(* IEC 61131-3 sources: 2026_Projet_YGO_ExcavatriceDragage/CODE/L_SIMULATION (part 2) *)

(* ---- FB_Sim_WinchElectrical.st ---- *)
(* ═══════════════════════════════════════════════════════════════
   🧪 FB_Sim_WinchElectrical — Composite electrique treuil (charge + couplage)
   ───────────────────────────────────────────────────────────────
   🎯 Role : Calcule le couple resistant reel (charge, benne au sol, couplage
   M1/M2) et pilote FB_Sim_WinchMotor. Transition de charge lissee (evite les
   a-coups de couple/vitesse a la bascule seul<->couple ou charge<->benne au sol).
   📄 Doc metier : DOC/WFLOW/CONTRACTS/PLAN_T317_SIMBENCH_TREUIL_ELECTRIQUE.md
   (registre sequence/interface 2026-09-18 -- pas encore integre a AF_Partie-13)
   🧩 Dependances : FB_Sim_WinchMotor
   ═══════════════════════════════════════════════════════════════ *)
FUNCTION_BLOCK PUBLIC FB_Sim_WinchElectrical
VAR_INPUT
    // === CONTRAT LIGHT ===
    Enable                    : BOOL; // --> [CMD] Autorisation generale FB

    // === COMMANDES ===
    StepCmd                   : INT;  // --> [CMD] Palier resistance rotorique actif (1..5)
    DirectionCmd              : INT := 1; // --> [CMD] Sens (1=Montee, -1=Descente)
    NetworkVoltageAct_V       : REAL := 400.0; // --> [HW] Tension reseau mesuree/simulee

    // === CHARGE ===
    LoadFrac_Ratio            : REAL; // --> [CMD] Taux de charge commande/estime (0..1)
    IsBucketGrounded          : BOOL; // --> [HW] TRUE = benne posee/cable detendu -> charge forcee a 0
        // A cabler sur l'image simulee de M2_TensionedCable_DI (NOT IsBucketGrounded) une fois le
        // stimulus expose en amont (GVL_Simulation) -- interface prete, cablage source en attente.
    LoadTransitionFilter_S    : REAL := 0.5; // --> [CFG] Constante de temps lissage charge (evite a-coup)

    // === COUPLAGE M1/M2 ===
    IsCoupledToPeer           : BOOL; // --> [CMD] TRUE = les deux treuils sont couples (benne commune)
        // A cabler sur l'equivalent simule de CoupledBoth/SyncActive (PRG_04_Treuils_Benne) une fois
        // expose en amont -- interface prete, cablage source en attente (lag 1 cycle accepte).
    PeerTorque_Nm             : REAL; // --> [BUS] Couple moteur de l'autre treuil (cycle precedent)
    PeerSpeed_Rpm             : REAL; // --> [BUS] Vitesse physique de l'autre treuil (cycle precedent)

    // === REGLAGES & CONFIGURATION (relayes a FB_Sim_WinchMotor) ===
    NetworkVoltageNom_V          : REAL := 400.0; // --> [CFG] Tension nominale reseau
    MaxTorque_Nm                 : REAL := 3800.0; // --> [CFG] Cmax decrochage -- SYNTHETIQUE
    SlipAtMaxTorqueBase_Ratio    : REAL := 0.08;   // --> [CFG] gmax palier rotor court-circuite
    RotorResistanceOwn_Ohm       : REAL := 0.08;   // --> [CFG] R2 propre rotor
    Inertia_KgM2                 : REAL := 45.0;   // --> [CFG] Inertie ramenee -- SYNTHETIQUE
    SynchronousSpeed_Rpm         : REAL := 1500.0; // --> [CFG] Vitesse synchronisme
    LoadNominalTorque_Nm         : REAL := 2500.0; // --> [CFG] Couple resistant a pleine charge -- SYNTHETIQUE
    LoadFrictionTorque_Nm        : REAL := 80.0;   // --> [CFG] Frottements residuels a vide -- SYNTHETIQUE
    CoupledPeerGain_Ratio         : REAL := 0.5;   // --> [CFG] Poids de l'effort differentiel du pair en mode couple
    CycleTime_S                  : REAL := 0.01;   // --> [CFG] Pas d'integration
END_VAR
VAR_OUTPUT
    // === CONTRAT LIGHT ===
    Ready                     : BOOL; // <-- [STAT] FB pret

    // === RESULTATS PHYSIQUES (relayes de FB_Sim_WinchMotor) ===
    MotorTorque_Nm            : REAL; // <-- [DIAG] Couple electromagnetique, repere de commande
    ResistiveTorqueAct_Nm     : REAL; // <-- [DIAG] Couple resistant reellement applique (charge+couplage, lisse)
    Slip_Ratio                : REAL; // <-- [DIAG] Glissement, repere de commande
    SpeedAct_Rpm               : REAL; // <-- [DIAG] Vitesse physique reelle signee (+montee/-descente)
    IsStalled                 : BOOL; // <-- [DIAG] Decrochage constate
    IsGeneratorMode            : BOOL; // <-- [DIAG] Mode freinage electrique
END_VAR
VAR
    // === SOUS-INSTANCE FB ===
    Motor                     : FB_Sim_WinchMotor; // * [INST] Couple electromagnetique elementaire

    // === ETAT INTERNE ===
    LoadFracFiltered_Ratio     : REAL; // . [LOC] Taux de charge lisse (PT1)
    LoadFracTarget_Ratio       : REAL; // . [LOC] Cible : 0 si benne au sol, sinon LoadFrac_Ratio
    PeerDifferentialTorque_Nm  : REAL; // . [LOC] Effort differentiel du pair en mode couple
    FilterAlpha_Ratio           : REAL; // . [LOC] Coefficient de lissage du pas courant
END_VAR
VAR CONSTANT
    CST_MinFilterTime_S        : REAL := 0.001;
END_VAR

// === §1 GATE NEUTRALISATION ===
IF NOT Enable THEN
    Ready := FALSE;
    MotorTorque_Nm := 0.0;
    ResistiveTorqueAct_Nm := 0.0;
    Slip_Ratio := 0.0;
    SpeedAct_Rpm := 0.0;
    IsStalled := FALSE;
    IsGeneratorMode := FALSE;
    LoadFracFiltered_Ratio := 0.0;
    RETURN;
END_IF;

// === §2 CHARGE LISSEE (benne au sol force la cible a 0, transition sans a-coup) ===
IF IsBucketGrounded THEN
    LoadFracTarget_Ratio := 0.0;
ELSE
    LoadFracTarget_Ratio := LIMIT(0.0, LoadFrac_Ratio, 1.0);
END_IF;

IF LoadTransitionFilter_S > CST_MinFilterTime_S THEN
    FilterAlpha_Ratio := CycleTime_S / (LoadTransitionFilter_S + CycleTime_S);
ELSE
    FilterAlpha_Ratio := 1.0;
END_IF;
LoadFracFiltered_Ratio := LoadFracFiltered_Ratio
    + FilterAlpha_Ratio * (LoadFracTarget_Ratio - LoadFracFiltered_Ratio);

// === §3 COUPLAGE M1/M2 ===
// En mode couple, la benne lie mecaniquement les deux treuils : un ecart de couple entre pairs
// se traduit en effort differentiel de rattrapage (proportionnel a l'ecart de vitesse), pas en
// deux dynamiques d'inertie totalement independantes qui divergent librement.
IF IsCoupledToPeer THEN
    PeerDifferentialTorque_Nm := CoupledPeerGain_Ratio * (SpeedAct_Rpm - PeerSpeed_Rpm)
        * LoadNominalTorque_Nm / MAX(SynchronousSpeed_Rpm, 1.0);
ELSE
    PeerDifferentialTorque_Nm := 0.0;
END_IF;

// === §4 COUPLE RESISTANT APPLIQUE ===
ResistiveTorqueAct_Nm := LoadFrictionTorque_Nm
    + DirectionCmd * LoadFracFiltered_Ratio * LoadNominalTorque_Nm
    + PeerDifferentialTorque_Nm;

// === §5 MOTEUR ELEMENTAIRE ===
Motor(
    Enable := TRUE,
    StepCmd := StepCmd,
    DirectionCmd := DirectionCmd,
    NetworkVoltageAct_V := NetworkVoltageAct_V,
    ResistiveTorque_Nm := ResistiveTorqueAct_Nm,
    NetworkVoltageNom_V := NetworkVoltageNom_V,
    MaxTorque_Nm := MaxTorque_Nm,
    SlipAtMaxTorqueBase_Ratio := SlipAtMaxTorqueBase_Ratio,
    RotorResistanceOwn_Ohm := RotorResistanceOwn_Ohm,
    Inertia_KgM2 := Inertia_KgM2,
    SynchronousSpeed_Rpm := SynchronousSpeed_Rpm,
    CycleTime_S := CycleTime_S
);

MotorTorque_Nm := Motor.MotorTorque_Nm;
Slip_Ratio := Motor.Slip_Ratio;
SpeedAct_Rpm := Motor.SpeedAct_Rpm;
IsStalled := Motor.IsStalled;
IsGeneratorMode := Motor.IsGeneratorMode;

Ready := TRUE;

(* ---- FB_Sim_WinchMotor.st ---- *)
(* ═══════════════════════════════════════════════════════════════
   🧪 FB_Sim_WinchMotor — Couple electromagnetique moteur treuil (rotor bobine)
   ───────────────────────────────────────────────────────────────
   🎯 Role : Couple (formule de Kloss), glissement bidirectionnel, decrochage
   predictif et mode generatrice pour un treuil M1/M2.
   📄 Doc metier : DOC/WFLOW/CONTRACTS/PLAN_T317_SIMBENCH_TREUIL_ELECTRIQUE.md
   (pas encore integre a AF_Partie-13 -- entree F13.06 a creer lot dedie)
   🧩 Dependances : FB_Sim_KlossTorque
   ═══════════════════════════════════════════════════════════════ *)
FUNCTION_BLOCK PUBLIC FB_Sim_WinchMotor
VAR_INPUT
    // === CONTRAT LIGHT ===
    Enable                    : BOOL; // --> [CMD] Autorisation generale FB (TRUE=Autorise)

    // === COMMANDES ===
    StepCmd                   : INT;  // --> [CMD] Palier resistance rotorique actif (1..5)
    DirectionCmd              : INT := 1; // --> [CMD] Sens (1=Montee, -1=Descente)

    // === MESURES / CHARGE ===
    NetworkVoltageAct_V       : REAL := 400.0; // --> [HW] Tension reseau mesuree/simulee
    ResistiveTorque_Nm        : REAL; // --> [CMD] Couple de charge DEJA projete en repere de
        // commande (N_rel) par l'appelant : positif = s'oppose au mouvement commande, negatif =
        // aide le mouvement (ex. gravite en descente -> peut declencher le mode generatrice).
        // Ce FB ne connait pas le taux de charge/la gravite -- calcul delegue a FB_Sim_WinchElectrical.

    // === REGLAGES & CONFIGURATION ===
    NetworkVoltageNom_V          : REAL := 400.0; // --> [CFG] Tension nominale reseau
    MaxTorque_Nm                 : REAL := 3800.0; // --> [CFG] Cmax decrochage -- SYNTHETIQUE
    SlipAtMaxTorqueBase_Ratio    : REAL := 0.08;   // --> [CFG] gmax au palier rotor court-circuite
        // (resistance externe nulle) -- SYNTHETIQUE. Sert de base a la mise a l'echelle par palier.
    RotorResistanceOwn_Ohm       : REAL := 0.08;   // --> [CFG] R2 propre rotor (palier court-circuite)
    Inertia_KgM2                 : REAL := 45.0;   // --> [CFG] Inertie ramenee -- SYNTHETIQUE
    SynchronousSpeed_Rpm         : REAL := 1500.0; // --> [CFG] Vitesse synchronisme
    CycleTime_S                  : REAL := 0.01;   // --> [CFG] Pas d'integration
END_VAR
VAR_OUTPUT
    // === CONTRAT LIGHT ===
    Ready                     : BOOL; // <-- [STAT] FB pret

    // === RESULTATS PHYSIQUES ===
    MotorTorque_Nm            : REAL; // <-- [DIAG] Couple electromagnetique, repere de commande
    Slip_Ratio                : REAL; // <-- [DIAG] Glissement, repere de commande
    SpeedAct_Rpm               : REAL; // <-- [DIAG] Vitesse physique reelle signee (+montee/-descente)
    IsStalled                 : BOOL; // <-- [DIAG] Decrochage constate (jamais reinitialise)
    IsGeneratorMode            : BOOL; // <-- [DIAG] Couple oppose au sens de commande (freinage)
END_VAR
VAR
    // === SOUS-INSTANCES FB ===
    KlossRunning               : FB_Sim_KlossTorque; // * [INST] Couple regime etabli
    KlossLockedRotor           : FB_Sim_KlossTorque; // * [INST] Couple test decrochage (g=1)

    // === ETAT INTERNE ===
    SpeedRel_RadPerS           : REAL; // . [LOC] Vitesse en repere de commande (N_rel)
    SynchronousSpeed_RadPerS   : REAL; // . [LOC] Vitesse synchronisme, rad/s
    SlipAtMaxTorqueStep_Ratio  : REAL; // . [LOC] gmax au palier courant
    SlipEff_Ratio               : REAL; // . [LOC] Glissement protege division par zero
    VoltageRatio2               : REAL; // . [LOC] (U_act/U_nom)^2
    Stalled                    : BOOL; // . [LOC] Etat instantane, peut se relever

    // === ENTREES BORNEES (SECURISE DIVISIONS) ===
    InertiaSafe_KgM2            : REAL; // . [LOC] Inertia_KgM2 bornee > 0
    RotorResistanceOwnSafe_Ohm  : REAL; // . [LOC] RotorResistanceOwn_Ohm bornee > 0
    SlipAtMaxTorqueBaseSafe_Ratio : REAL; // . [LOC] SlipAtMaxTorqueBase_Ratio bornee > 0
    NetworkVoltageNomSafe_V     : REAL; // . [LOC] NetworkVoltageNom_V bornee > 0
    StepCmdSafe                : INT;  // . [LOC] StepCmd borne [1..5]
END_VAR
VAR CONSTANT
    CST_StepCount              : INT := 5;
    CST_RotorExtResistanceStep_Ohm : ARRAY[1..5] OF REAL := [3.6, 1.9, 0.9, 0.35, 0.0];
        // palier 1 = resistance max (demarrage), palier 5 = rotor court-circuite -- SYNTHETIQUE
        // (indexation/valeurs propres au ST, pas un portage 1:1 du prototype Python 4 gradins)
    CST_MinSlip_Ratio          : REAL := 0.0001;
    CST_MinDenominator         : REAL := 0.001; // plancher generique config sensible (division)
    CST_StallSpeedThreshold_Rpm : REAL := 28.0; // ~3 rad/s, "quasi arrete"
END_VAR

// === §1 GATE NEUTRALISATION ===
IF NOT Enable THEN
    Ready := FALSE;
    MotorTorque_Nm := 0.0;
    Slip_Ratio := 0.0;
    SpeedAct_Rpm := 0.0;
    IsStalled := FALSE;
    IsGeneratorMode := FALSE;
    SpeedRel_RadPerS := 0.0;
    RETURN;
END_IF;

StepCmdSafe := LIMIT(1, StepCmd, CST_StepCount);
IF StepCmdSafe <> StepCmd THEN
    Ready := FALSE;
    RETURN;
END_IF;
IF (DirectionCmd <> 1) AND (DirectionCmd <> -1) THEN
    Ready := FALSE;
    RETURN;
END_IF;

// Bornage systematique des entrees de config sensibles (denominateurs) -- CODE_QUALITY_STANDARDS §6
InertiaSafe_KgM2 := MAX(CST_MinDenominator, Inertia_KgM2);
RotorResistanceOwnSafe_Ohm := MAX(CST_MinDenominator, RotorResistanceOwn_Ohm);
SlipAtMaxTorqueBaseSafe_Ratio := MAX(CST_MinDenominator, SlipAtMaxTorqueBase_Ratio);
NetworkVoltageNomSafe_V := MAX(1.0, NetworkVoltageNom_V);

// === §2 GLISSEMENT ET COUPLE (FORMULE DE KLOSS) ===
SynchronousSpeed_RadPerS := SynchronousSpeed_Rpm * 2.0 * 3.14159265 / 60.0;

// gmax(palier) = gmax_base * R2_total(palier) / R2_rotor_propre -- ajouter de la resistance
// externe deplace le glissement au couple max vers 1 (couple demarrage), sans changer Cmax.
// gmax_base = gmax au palier rotor court-circuite (resistance externe nulle).
SlipAtMaxTorqueStep_Ratio := SlipAtMaxTorqueBaseSafe_Ratio
    * (RotorResistanceOwnSafe_Ohm + CST_RotorExtResistanceStep_Ohm[StepCmdSafe])
    / RotorResistanceOwnSafe_Ohm;

// Glissement en repere de commande (N_rel) : peut etre negatif (survitesse -> freinage
// generateur). SpeedRel_RadPerS reste dans ce repere ; SpeedAct_Rpm restitue le signe physique.
Slip_Ratio := 1.0 - SpeedRel_RadPerS / SynchronousSpeed_RadPerS;

IF ABS(Slip_Ratio) < CST_MinSlip_Ratio THEN
    IF Slip_Ratio >= 0.0 THEN
        SlipEff_Ratio := CST_MinSlip_Ratio;
    ELSE
        SlipEff_Ratio := -CST_MinSlip_Ratio;
    END_IF;
ELSE
    SlipEff_Ratio := Slip_Ratio;
END_IF;

VoltageRatio2 := (NetworkVoltageAct_V / NetworkVoltageNomSafe_V) * (NetworkVoltageAct_V / NetworkVoltageNomSafe_V);

KlossRunning(
    Enable := TRUE,
    MaxTorque_Nm := MaxTorque_Nm,
    Slip_Ratio := SlipEff_Ratio,
    SlipAtMaxTorque_Ratio := SlipAtMaxTorqueStep_Ratio,
    VoltageRatio2 := VoltageRatio2);
MotorTorque_Nm := KlossRunning.Torque_Nm;

// === §3 DYNAMIQUE MECANIQUE ===
// Pas de saturation basse : SpeedRel_RadPerS peut devenir negatif (glissement arriere sous
// surcharge) ou depasser le synchronisme (regime generateur).
SpeedRel_RadPerS := SpeedRel_RadPerS
    + (MotorTorque_Nm - ResistiveTorque_Nm) / InertiaSafe_KgM2 * CycleTime_S;

SpeedAct_Rpm := SpeedRel_RadPerS * DirectionCmd * 60.0 / (2.0 * 3.14159265);

// === §4 DECROCHAGE PREDICTIF ===
// Au palier courant, couple disponible a glissement bloque (g=1) < couple resistant, ET
// vitesse quasi nulle -- prediction "ce palier peut-il tenir la charge depuis l'arret ?",
// pas une mesure d'arret reel.
IF ABS(SpeedAct_Rpm) < CST_StallSpeedThreshold_Rpm THEN
    KlossLockedRotor(
        Enable := TRUE,
        MaxTorque_Nm := MaxTorque_Nm,
        Slip_Ratio := 1.0,
        SlipAtMaxTorque_Ratio := SlipAtMaxTorqueStep_Ratio,
        VoltageRatio2 := VoltageRatio2);
    Stalled := KlossLockedRotor.Torque_Nm < ResistiveTorque_Nm;
    IF Stalled THEN
        IsStalled := TRUE;
    END_IF;
ELSE
    Stalled := FALSE;
END_IF;

IsGeneratorMode := MotorTorque_Nm < 0.0;

Ready := TRUE;

(* ---- FB_SimBench.st ---- *)
(* ═══════════════════════════════════════════════════════════════
   🧪 FB_SimBench — Enveloppe unique de simulation pour banc d'essai
   ───────────────────────────────────────────────────────────────
   📄 Doc métier : DOC/AF/AF_Partie-13_Fonction_Simulation_v2.5.md

   🎯 Rôle : Compose les blocs de modèle de simulation :
      - FB_Sim_Encoder (instM1, instM2)
      - FB_Sim_Translation (instTranslation)
      - FB_Sim_Joystick (instJoystick)
      - FB_Sim_Safety (instSafety)

   🔒 Brique réduite : 0 lecture de variable globale en interne.
      Toutes les entrées (commandes, stimuli, HwReal) sont passées en paramètres.

   🔴 RÈGLES SÉCURITÉ ET POLARITÉ :
      - Modèle frein M1/M2/M3 : M1_BrakeIsOpen_DI := M1_BrakeCmd (1 = OUVERT).
        Ne JAMAIS faire NOT BrakeCmd !
      - Retours contacteurs M1/M2 : 1 = tous retombés (TRUE quand RelayFwd=0 et RelayRev=0).
   ═══════════════════════════════════════════════════════════════ *)

FUNCTION_BLOCK PUBLIC FB_SimBench
VAR_INPUT
    Enable                     : BOOL;             (* --> [CMD] Activation globale (GVL_Simulation.SimulationModeActive) *)
    OperatorSourceActive       : BOOL := TRUE;      (* --> [CMD] Source operateur simulee effectivement selectionnee *)

    // ── Commandes issues de l'automate (Scan N-1 / PRG_07 / PRG_10) ──────────
    M1_RelayFwd                : BOOL;   (* --> [CMD] Sens avant M1 *)
    M1_RelayRev                : BOOL;   (* --> [CMD] Sens arrière M1 *)
    // Les 4 contacteurs de palier participent au retour unique
    // « tous contacteurs retombés » — sans eux, le modèle annonce l'arrêt alors qu'un
    // palier est encore engagé (fausse condition d'armement Méca A).
    M1_SpeedContactor_1        : BOOL;   (* --> [HW] Contacteur palier 1 M1 *)
    M1_SpeedContactor_2        : BOOL;   (* --> [HW] Contacteur palier 2 M1 *)
    M1_SpeedContactor_3        : BOOL;   (* --> [HW] Contacteur palier 3 M1 *)
    M1_SpeedContactor_4        : BOOL;   (* --> [HW] Contacteur palier 4 M1 *)
    M1_SpeedCmd_Pct            : REAL;   (* --> [CMD] Consigne vitesse M1 *)
    M1_StepNumber              : INT;    (* --> [CMD] Palier vitesse courant M1 (1..5) *)
    M1_PresetTriggerCmd        : WORD;   (* --> [CMD] Trigger preset M1 *)
    M1_PresetValueOut          : UDINT;   (* --> [CFG] Valeur preset M1 *)
    M1_BrakeCmd                : BOOL;             (* --> [CMD] TRUE = commande desserrage frein M1 *)

    M2_RelayFwd                : BOOL;   (* --> [CMD] Sens avant M2 *)
    M2_RelayRev                : BOOL;   (* --> [CMD] Sens arrière M2 *)
    M2_SpeedContactor_1        : BOOL;   (* --> [HW] Idem M1, voir ci-dessus *)
    M2_SpeedContactor_2        : BOOL;   (* --> [HW] Contacteur palier 2 M2 *)
    M2_SpeedContactor_3        : BOOL;   (* --> [HW] Contacteur palier 3 M2 *)
    M2_SpeedContactor_4        : BOOL;   (* --> [HW] Contacteur palier 4 M2 *)
    M2_SpeedCmd_Pct            : REAL;   (* --> [CMD] Consigne vitesse M2 *)
    M2_StepNumber              : INT;    (* --> [CMD] Palier vitesse courant M2 (1..5) *)
    M2_PresetTriggerCmd        : WORD;   (* --> [CMD] Trigger preset M2 *)
    M2_PresetValueOut          : UDINT;   (* --> [CFG] Valeur preset M2 *)
    M2_BrakeCmd                : BOOL;             (* --> [CMD] TRUE = commande desserrage frein M2 *)

    M3_ReqTremie               : BOOL;             (* --> [CMD] Demande explicite vers Trémie *)
    M3_ReqMaintenance          : BOOL;             (* --> [CMD] Demande explicite vers Maintenance *)
    M3_SpeedCmd_Pct            : REAL;   (* --> [CMD] Consigne vitesse M3 *)
    (* T301/L1 — SOURCE UNIQUE : reglages machine M3 lus par PRG_02 (le banc n'a plus de positions en dur) *)
    M3_PosTremie_M             : REAL := 0.0;   (* --> [CFG] Position capteur Tremie (GVL_PERSISTENT) *)
    M3_PosPV_M                 : REAL := 1.5;   (* --> [CFG] Position capteur PV (GVL_PERSISTENT) *)
    M3_PosP2_M                 : REAL := 3.5;   (* --> [CFG] Position capteur P2 (GVL_PERSISTENT) *)
    M3_PosP1_M                 : REAL := 5.0;   (* --> [CFG] Position capteur P1 (GVL_PERSISTENT) *)
    M3_PosMaintenance_M        : REAL := 10.0;  (* --> [CFG] Position capteur Maintenance (GVL_PERSISTENT) *)
    M3_OdometryGain            : REAL := 0.02;  (* --> [CFG] Gain effectif de l'estimateur machine, m/(Hz.s) (PRG_05) *)
    M3_EstimatedPos_M          : REAL;          (* --> [DIAG] Position calculee par le programme (PRG_05), pour l'ecart observe *)
    M3_BrakeCmd                : BOOL;             (* --> [CMD] TRUE = commande desserrage frein M3 *)

    PowerKeepAlive_A           : BOOL;             (* --> [SAFE] TRUE = relais A maintenu sagement par le PLC *)
    PowerKeepAlive_B           : BOOL;             (* --> [SAFE] TRUE = relais B maintenu sagement par le PLC *)
    EmergencyArming_RQ         : BOOL;             (* --> [CMD] Impulsion de réarmement puissance *)
    TestCutActive              : BOOL;             (* --> [SAFE] Test de redondance AU en cours (canal A ou B coupé) *)
    PowerCutOffRequest         : BOOL;             (* --> [SAFE] Requête coupure métier (TRUE = arrêt d'urgence) *)
    SimChainOkBit              : BOOL;             (* --> [TST] Bit opérateur : TRUE = simuler chaîne AU fermée *)
    SimPhaseRotationOkBit      : BOOL;             (* --> [TST] Bit opérateur : TRUE = phases réseau OK ; FALSE = défaut rotation de phases *)

    // ── Stimuli & Paramètres de banc ─────────────────────────────────────────
    SimEncoderSpeedFactor      : REAL := 1.0;   (* --> [CFG] Facteur vitesse codeur *)
    SimBucketSpeedFactor       : REAL := 1.0;   (* --> [CFG] Facteur vitesse manoeuvre benne seule (non persistant) *)
    SimTopPositionActive       : BOOL := FALSE; (* --> [TST] Injection manuelle capteur haut actif (essai ciblé) *)
    SimSyncDeviationInjectM1   : BOOL := FALSE;   (* --> [TST] Injection écart synchro M1 *)
    SimSyncDeviationInjectM2   : BOOL := FALSE;   (* --> [TST] Injection écart synchro M2 *)
    SimSyncDeviationOffset_M   : REAL := 0.5;   (* --> [TST] Offset écart synchro *)
    SimM2CoupledDescentModelActive : BOOL := TRUE; (* --> [CFG] M2 calculé depuis M1 en descente BOTH *)
    SimM2CoupledDescentFactor  : REAL := 0.9333; (* --> [CFG] Ratio déplacement M2/M1 mesuré: 0,6m d'écart sur 9m *)
    SimWinchSpeedReportTauS    : REAL := 0.0;    (* --> [CFG][SYNTHETIQUE] Tau 1er ordre retour vitesse rapportee M1/M2, s. 0.0 = saut instantane (comportement historique). *)
    SimWinchBrakeOpenDelayS    : REAL := 0.0;    (* --> [CFG][SYNTHETIQUE] Delai electrique/meca ouverture frein M1/M2 apres BrakeCmd=TRUE, s. 0.0 = instantane (comportement historique). *)
    SimWinchBrakeCloseDelayS   : REAL := 0.0;    (* --> [CFG][SYNTHETIQUE] Delai electrique/meca fermeture frein M1/M2 apres BrakeCmd=FALSE, s. 0.0 = instantane (comportement historique). *)
    SimWinchDynamicsActive     : BOOL := FALSE;  (* --> [CFG] TRUE = applique tau et delais treuils ; FALSE = profil simple historique *)

    // T317 exploratoire -- charge/couplage electrique treuil (interface prete, defaut = comportement
    // historique inchange tant que non cablee sur un vrai signal amont, cf. registre PLAN_T317).
    SimWinchLoadFrac_Ratio     : REAL := 0.0;    (* --> [CFG][SYNTHETIQUE] Taux de charge M1/M2, 0=a vide *)
    SimWinchCoupledActive      : BOOL := FALSE;  (* --> [TST] M1/M2 couples -- en attente cablage CoupledBoth reel *)
    SimWinchElectricalDiagnosticsActive : BOOL := FALSE; (* --> [CFG] TRUE = publie diagnostic electrique treuils, sans action safety *)
    SimM2TensionedCableFaultInject : BOOL := FALSE; (* --> [TST] TRUE = injecte capteur cable non tendu M2 *)

    SimM3SensorsWordOverrideActive : BOOL := FALSE;   (* --> [TST] Override mot capteurs M3 *)
    SimM3SensorsWord               : BYTE := 16#07;   (* --> [TST] Mot capteurs M3 forcé *)
    SimM3SensorIntermittenceActive  : BOOL := FALSE;   (* --> [TST] Episode perte/reprise DI M3 *)
    SimM3SensorStabilizationS       : REAL := 1.0;     (* --> [CFG] Duree episode capteur M3, s *)
    SimM3SensorElectricalDelayS     : REAL := 0.01;    (* --> [CFG] Delai electrique capteur M3, s *)
    SimM3SensorIntermittencePeriodS : REAL := 0.12;    (* --> [CFG] Periode des bascules episode, s *)
    SimM3SensorHysteresis_M         : REAL := 0.02;    (* --> [CFG] Hysteresis seuils capteurs M3, m *)
    SimM3SensorLoadAngleTriggerRad  : REAL := 0.01;    (* --> [CFG] Angle charge minimal episode, rad *)
    SimM3SensorScenarioSeed         : UDINT := 3001;   (* --> [CFG] Graine episode capteurs M3 *)
    SimM3SensorBlipTransitions      : UDINT := 0;      (* --> [TST] Excursions electriques courtes par front (0 = profil ~1 s historique seul) *)
    SimM3SensorBlipDurationS        : REAL := 0.2;     (* --> [CFG] Largeur d'une excursion du blip court, s *)
    // FAUTE explicite frein M3 — defaut FALSE : reproduit le defaut terrain « frein ferme
    // alors que le variateur retourne encore 10,00 Hz » (trace 2026-09-04, 26,437 s, ErrorId=64).
    SimM3BrakeFaultCloseWhileRunning : BOOL := FALSE;  (* --> [TST] TRUE = force la fermeture frein M3 hors vitesse nulle *)
    SimM3BrakeFaultCloseDelayS       : REAL := 0.0;    (* --> [CFG] Delai avant application de la faute frein M3, s *)
    SimM3BrakePhysicalActive         : BOOL := TRUE;   (* --> [CFG] L3 : frein M3 a manque de courant reel (FALSE = historique) *)
    SimM3BrakeDecel_Mps2             : REAL := 2.0;    (* --> [CFG][HYPOTHESE] Deceleration chariot frein serre, m/s2 *)
    SimM3CartFreeActive              : BOOL := TRUE;   (* --> [CFG] L4 : chariot libre frein ouvert + variateur sans couple *)
    SimM3LoadMassRatio               : REAL := 0.5;    (* --> [CFG][HYPOTHESE] Masse benne / masse totale *)
    SimM3RollingFriction_Mps2        : REAL := 0.1;    (* --> [CFG][HYPOTHESE] Frottement de roulement, m/s2 *)
    SimM3Slope_Mps2                  : REAL := 0.0;    (* --> [CFG][HYPOTHESE] Pente, m/s2 (+ vers Maintenance) *)
    SimM3SensorCamDropoutActive      : BOOL := TRUE;   (* --> [CFG] L5 : came capteurs vu -> perdu -> retrouve -> fixe *)
    SimM3SensorCamDropoutStart_M     : REAL := 0.02;   (* --> [CFG][HYPOTHESE] Debut de la zone perdue apres la cote, m *)
    SimM3SensorCamDropoutWidth_M     : REAL := 0.04;   (* --> [CFG][HYPOTHESE] Largeur de la zone perdue, m *)
    // BUTEE MECANIQUE M3 — recul borne apres arret serre (C5). 0.0 = comportement historique
    // (position ET vitesse figees a la butee, decision de review tracee). > 0 autorise la
    // reaction de charge a ressortir le chariot de la zone capteur. SYNTHETIQUE, non calibre.
    SimM3EndStopRecoilMax_M          : REAL := 0.0;    (* --> [CFG][SYNTHETIQUE] Recul borne a la butee M3, m *)
    SimM3EndStopMargin_M             : REAL := 0.5;    (* --> [CFG] Distance capteur extreme -> butee mecanique M3, m *)
    SimM3LoadReactionGain_Mps2       : REAL := 0.20;   (* --> [CFG][SYNTHETIQUE] Gain de reaction de charge M3, m/s2 *)
    // ACCELERATION DU BANC M3 : chariot ET frequence retournee x facteur (1..5), estimation coherente.
    // Volontairement NON cable par PRG_02 : se regle en ligne sur l'instance (instSimBench.SimM3SpeedFactor).
    SimM3SpeedFactor                 : REAL := 1.0;    (* --> [TST] Facteur de vitesse du banc M3, 1,0 = dynamique reelle *)

    SimJoystickLeft_Rev_TREMIE_Active  : BOOL := FALSE;   (* --> [TST] Bouton joystick gauche *)
    SimJoystickRight_Fwd_MAINT_Active  : BOOL := FALSE;   (* --> [TST] Bouton joystick droite *)
    SimJoystickFwd_Up_Close_Active     : BOOL := FALSE;   (* --> [TST] Bouton joystick avant *)
    SimJoystickRev_Down_Open_Active    : BOOL := FALSE;   (* --> [TST] Bouton joystick arrière *)
    SimJoystickRawX                    : INT := 5000;   (* --> [TST] Valeur brute X *)
    SimJoystickRawY                    : INT := 5000;   (* --> [TST] Valeur brute Y *)
    SimJoystickRawButton               : BOOL := FALSE;   (* --> [TST] Bouton homme-mort *)
    SimJoystickOvershoot_Active        : BOOL := FALSE;   (* --> [TST] Dépassement de montée au-delà de 100% (défaut capteur hors plage) *)
    SimJoystickBagotement_Active       : BOOL := FALSE;   (* --> [TST] Bagotement au relâchement (petit balancement autour du neutre) *)

    SimKoboldContactValue      : BOOL := FALSE;   (* --> [TST] Contact fond Kobold *)
    SimKoboldAutoModeActive    : BOOL := FALSE;   (* --> [CFG] Kobold positionnel automatique armé *)
    SimKoboldAutoDepth_M       : REAL := -15.0;   (* --> [CFG] Fond Kobold signé *)
    SimKoboldPowerUpTime       : TIME := T#50ms;  (* --> [CFG] Temps de réponse sonde *)
    SimKoboldCoast_M           : REAL := 1.0;     (* --> [CFG] Compatibilité interface ; dynamique historique utilisée *)
    KoboldMeasureEnable        : BOOL := FALSE;   (* --> [CMD] Alimentation Kobold effectivement arbitrée *)
    M1_CablePos_M              : REAL := 0.0;     (* --> [HW] Position M1 signée, référence homing effective *)
    BtnEmergencyStop           : BOOL := FALSE;    (* --> [TST] Simulation appui coup-de-poing AU *)

    // ── Rattrapage mécanique M1/M2 (reprise de jeu en mouvement couplé) ──
    SimWinchCouplingModelActive : BOOL := TRUE;    (* --> [CFG] TRUE = rattrapage mécanique modélisé au banc *)
    SimBucketJamActive          : BOOL := FALSE;   (* --> [TST] TRUE = mâchoires bloquées (objet coincé) *)
    WinchesHomed                : BOOL := TRUE;    (* --> [HW] TRUE = M1 et M2 references (butee meca benne inactive avant homing) *)
    M2_CablePos_M               : REAL := 0.0;     (* --> [HW] Position M2 recalée (m), issue de la même chaîne que le métier *)
    BucketOffsetCloseM          : REAL := 15.0;    (* --> [CFG] Butée mécanique benne FERMÉE (m, écart M2-M1) *)
    BucketCoherenceLimitM       : REAL := 1.0;     (* --> [CFG] Demi-largeur de la bande franc ouvert/fermé (m) *)
    BucketOffsetOpen_M          : REAL := 0.0;     (* --> [CFG] Butée mécanique benne OUVERTE (m, écart M2-M1) *)
    BucketOpenAnticipation_M    : REAL := 1.3;     (* --> [CFG] Anticipation arrêt ouverture benne (m) *)
    BucketAx15bOpenActive       : BOOL := FALSE;   (* --> [CMD] Étape AX15B active *)

    // ── Image réelle fallback ────────────────────────────────────────────────
    HwReal                     : ST_HardwareImage;   (* --> [HW] Image réelle fallback *)
END_VAR

VAR_OUTPUT
    (* Sorties d'état du profil AF_Partie-03 §2.
       En LD, CODESYS réserve la PREMIÈRE broche de sortie au flux du rung :
       `Ready` n'y porte jamais d'expression, les broches suivantes oui. *)
    Ready                      : BOOL;             (* <-- [STAT] TRUE = banc prêt (Enable actif, modèles à jour) *)
    Busy                       : BOOL;             (* <-- [STAT] TRUE = cycle de simulation en cours *)
    Done                       : BOOL;             (* <-- [STAT] TRUE = images de simulation publiées ce scan *)

    Winch                      : ST_HwWinch;   (* <-- [DIAG] Image treuils simulée *)
    Translation                : ST_HwTranslation;   (* <-- [DIAG] Image translation simulée *)
    Operator                   : ST_HwOperator;   (* <-- [DIAG] Image opérateur simulée *)
    Machine                    : ST_HwMachine;   (* <-- [DIAG] Image machine simulée *)

    // T317 exploratoire -- modele electrique treuil, diagnostic seul, non consomme par le metier.
    // Charge appliquee = LoadFrictionTorque_Nm + taux x LoadNominalTorque_Nm (FB_Sim_WinchElectrical) ;
    // le taux de charge n'est pas encore cable sur un signal amont (registre PLAN_T317).
    MotorTorqueM1_Nm           : REAL;   (* <-- [DIAG] T317 -- Couple electromagnetique simule M1 *)
    MotorTorqueM2_Nm           : REAL;   (* <-- [DIAG] T317 -- Couple electromagnetique simule M2 *)
    MotorIsStalledM1           : BOOL;   (* <-- [DIAG] T317 -- Decrochage predictif simule M1 *)
    MotorIsStalledM2           : BOOL;   (* <-- [DIAG] T317 -- Decrochage predictif simule M2 *)

    // Rattrapage mecanique M1/M2 -- diagnostic seul (aucun consommateur metier).
    WinchCouplingActive        : BOOL;   (* <-- [DIAG] Rattrapage applique ce scan *)
    WinchCouplingCorrectionPts : DINT;   (* <-- [DIAG] Correction appliquee a l'image M2 (points codeur) *)

    // Faute frein M3 -- diagnostic seul : confirme que la branche de faute est bien appliquee.
    M3BrakeFaultCloseActive    : BOOL;   (* <-- [DIAG] Faute frein M3 effectivement appliquee ce scan *)
    // Blip court capteurs M3 -- diagnostic seul : observable sur trace pendant un episode court.
    M3SensorBlipActive         : BOOL;   (* <-- [DIAG] Un capteur M3 publie une excursion courte *)
    (* L2 — observation M3 (lecture seule, aucun effet sur le pilotage) *)
    M3ObsPositionTrue_M        : REAL;   (* <-- [DIAG] Position vraie du chariot simule (m) *)
    M3ObsPositionError_M       : REAL;   (* <-- [DIAG] Position vraie - position calculee par le programme (m) *)
    M3ObsOvershootLast_M       : REAL;   (* <-- [DIAG] Distance roulee apres le 1er front du dernier capteur d'arret (m) *)
    M3ObsOvershootSensorId     : INT;    (* <-- [DIAG] 1 = Tremie, 3 = P1, 5 = Maintenance *)
    M3ObsEndStopHitCount       : UDINT;  (* <-- [DIAG] Chocs en butee mecanique *)
    M3ObsEndStopImpactSpeed_Mps : REAL;  (* <-- [DIAG] Vitesse au dernier choc en butee (m/s) *)
    M3ObsBrakeClosedMovingCount : UDINT; (* <-- [DIAG] Fermetures du frein chariot en mouvement *)
    M3ObsCartFree              : BOOL;   (* <-- [DIAG] L4 : chariot libre (frein ouvert, variateur sans couple) *)
    M3ObsFreeRollLast_M        : REAL;   (* <-- [DIAG] L4 : distance du dernier episode libre (m) *)
END_VAR

VAR_IN_OUT
    // 🔒 LECTURE SEULE pour le banc : ces mémoires appartiennent au modèle codeur. Le banc les lit
    //    pour piloter ses modèles et ne les écrit JAMAIS — pas même pour « initialiser » une mémoire
    //    lue à 0 (un 0 est un point de passage légitime du comptage signé, jamais une mémoire vierge).
    RawPosM1                   : UDINT;            (* <-> [BUS] Mémoire _SimEncoderRawPosM1 dans GVL_PERSISTENT *)
    RawPosM2                   : UDINT;            (* <-> [BUS] Mémoire _SimEncoderRawPosM2 dans GVL_PERSISTENT *)
END_VAR

VAR CONSTANT
    // T301/L1 : l'ancienne echelle en dur CST_M3FullTravelTimeS (37,5 s) est SUPPRIMEE — le banc
    // recoit positions + gain effectif de la machine (M3_Pos*_M, M3_OdometryGain). Gate G518.
    // Maximum variateur M3 : DOIT egaler GVL_PERSISTENT._TranslationMaxFreq_Hz (PRG_02 envoie f/50 x 100).
    // Constante locale (L_SIMULATION ne lit pas GVL_PERSISTENT) ; egalite verifiee par G518.
    CST_M3MaxFreq_Hz            : REAL := 50.0;
    CST_SimBenchCycleTimeS      : REAL := 0.010; // Période tâche PLC (s) — MainTask 10 ms
    // Rattrapage mécanique M1/M2 — valeurs ESTIMÉES (voir REGISTRE_VALEURS_TREUIL_STATUTS_v1.0.md)
    CST_SimWinchCouplingTauS    : REAL := 1.0;   // [HYPOTHESE] Constante de temps du rattrapage (s)
    CST_SimWinchCouplingStepMax_M : REAL := 0.02; // [HYPOTHESE] Borne de pente par scan (= 2,0 m/s x 0,010 s)
    CST_SimWinchCouplingPtsPerM : REAL := 4096.0; // Points codeur par mètre (8192 pts/tour / 2,0 m/tour)
    CST_SimBucketJamLoadFrac_Ratio : REAL := 1.0; // [HYPOTHESE] Charge forcée quand les mâchoires sont bloquées
END_VAR

VAR
    // Modèles sous-jacents
    instSimEncoderM1           : FB_Sim_Encoder;   (* * [INST] Modèle codeur M1 *)
    instSimEncoderM2           : FB_Sim_Encoder;   (* * [INST] Modèle codeur M2 *)
    instSimTranslation         : FB_Sim_Translation;   (* * [INST] Modèle translation M3 *)
    instSimJoystick            : FB_Sim_Joystick;   (* * [INST] Modèle joystick *)
    instSimSafety              : FB_Sim_Safety;   (* * [INST] Modèle sécurité *)
    instWinchElectricalM1      : FB_Sim_WinchElectrical;   (* * [INST] T317 exploratoire -- electrique+charge M1 *)
    instWinchElectricalM2      : FB_Sim_WinchElectrical;   (* * [INST] T317 exploratoire -- electrique+charge M2 *)
    PeerTorqueM1Prev_Nm        : REAL;   (* . [LOC] T317 -- couple M1 cycle precedent, pour M2 couple *)
    PeerTorqueM2Prev_Nm        : REAL;   (* . [LOC] T317 -- couple M2 cycle precedent, pour M1 couple *)
    PeerSpeedM1Prev_Rpm        : REAL;   (* . [LOC] T317 -- vitesse M1 cycle precedent, pour M2 couple *)
    PeerSpeedM2Prev_Rpm        : REAL;   (* . [LOC] T317 -- vitesse M2 cycle precedent, pour M1 couple *)
    KoboldBottomTouchPrev_DI   : BOOL;   (* . [LOC] T317 -- Machine.M1_M2_KoboldBottomTouch_DI cycle precedent (benne au sol) *)

    // Calculs internes
    M1_PresetCmd               : BOOL;   (* . [LOC] Trigger preset M1 *)
    M2_PresetCmd               : BOOL;   (* . [LOC] Trigger preset M2 *)
    M1_OffsetPts               : DINT;   (* . [LOC] Offset synchro M1 *)
    M2_OffsetPts               : DINT;   (* . [LOC] Offset synchro M2 *)

    M3_RelayFwd                : BOOL;   (* . [LOC] Sens avant M3 *)
    M3_RelayRev                : BOOL;   (* . [LOC] Sens arrière M3 *)

    SimJoystickManualNeutral : BOOL; (* . [LOC] Axes manuels au neutre nominal *)
    SimJoystickGesturePermit : BOOL; (* . [LOC] Aucune injection manuelle concurrente au geste *)

    M3_ActualFreqHz            : UINT;   (* . [LOC] Fréquence simulée M3 *)
    M3_StatusWordSim           : WORD;   (* . [LOC] StatusWord simulé M3 *)

    // Roulis dynamique avec dispersion pseudo-aléatoire (±0.1m autour de l'anticipation)
    M2_RelayFwdPrev            : BOOL;   (* . [LOC] Mémoire relais Fwd N-1 *)
    M2_RelayRevPrev            : BOOL;   (* . [LOC] Mémoire relais Rev N-1 *)
    RandomSeed                 : UDINT := 123456789; (* . [LOC] Générateur LCG pseudo-aléatoire *)
    M2_EffectiveCoastM         : REAL := 1.30;       (* . [LOC] Distance de roulis M2 courante *)
    M2EffectiveCoastDistance_M : REAL;               (* . [LOC] Distance appliquée au codeur M2 *)
    M2AutoOpenCoastArmed       : BOOL;               (* . [LOC] Fin d'ouverture automatique à simuler *)
    M2OpenDistanceRemaining_M  : REAL;               (* . [LOC] Distance restante à la butée ouverte *)
    M2OpenStopThreshold_M     : REAL;               (* . [LOC] Seuil avec avance d'un scan d'acquisition *)
    M2ExpectedStepDistance_M  : REAL;               (* . [LOC] Course codeur M2 du scan actif *)
    M2BucketOnlyActive         : BOOL;                (* . [LOC] Manœuvre benne seule (M2 actif, M1 au repos) *)
    SpeedM1_Mps                : REAL;                (* . [LOC] Vitesse nominale palier M1 m/s *)
    SpeedM2_Mps                : REAL;                (* . [LOC] Vitesse nominale palier M2 m/s *)
    M2CoupledDescentActive     : BOOL;                (* . [LOC] Ralentissement M2 actif en descente BOTH *)
    M2_MechanicStopEngaged     : BOOL;                (* . [LOC] Butee mecanique benne atteinte (T421) *)
    M2EffectiveSpeedScaleFactor : REAL;               (* . [LOC] Facteur vitesse du producteur unique M2 *)
    KoboldMeasureEnablePrevious : BOOL;               (* . [LOC] Front alimentation Kobold *)

    // Rattrapage mecanique M1/M2 : reprise de jeu entre les deux treuils
    WinchCouplingBothSameDir   : BOOL;   (* . [LOC] Les deux relais de sens actifs dans le meme sens *)
    WinchCouplingGate          : BOOL;   (* . [LOC] Condition complete de rattrapage *)
    WinchCouplingDelta_M       : REAL;   (* . [LOC] Ecart relatif M2-M1 courant (m) *)
    WinchCouplingCorrection_M  : REAL;   (* . [LOC] Correction calculee ce scan (m) *)
    WinchCouplingCorrectionDInt : DINT;  (* . [LOC] Correction convertie en points codeur *)
    WinchCouplingTarget_M      : REAL;   (* . [LOC] Entree de bande fermee visee (m) *)
    WinchCouplingAccumPts      : DINT;   (* . [LOC] Reprise de jeu accumulee sur l'image M2 (points) *)
    KoboldAutoEpisodeActive    : BOOL;                (* . [LOC] Mode auto figé pour une plongée *)
    KoboldAutoDepthEpisode_M   : REAL;                (* . [LOC] Fond figé durant une plongée *)
    KoboldPowerUpEpisodeTime   : TIME;                (* . [LOC] Délai sonde figé durant une plongée *)
    instKoboldPowerUpTimer     : TON;                 (* . [LOC] Réponse sonde après alimentation *)

    // Dynamique treuil M1/M2 : delais opt-in — defaut 0.0 = comportement historique
    M1_BrakeIsOpenState        : BOOL;                (* . [LOC] Etat frein M1 filtre par le delai *)
    M1_BrakeOpenTimerS         : REAL;                (* . [LOC] Accumulateur delai ouverture frein M1 *)
    M1_BrakeCloseTimerS        : REAL;                (* . [LOC] Accumulateur delai fermeture frein M1 *)
    M2_BrakeIsOpenState        : BOOL;                (* . [LOC] Etat frein M2 filtre par le delai *)
    M2_BrakeOpenTimerS         : REAL;                (* . [LOC] Accumulateur delai ouverture frein M2 *)
    M2_BrakeCloseTimerS        : REAL;                (* . [LOC] Accumulateur delai fermeture frein M2 *)
    WinchSpeedReportTauEffectiveS : REAL;             (* . [LOC] Tau applique apres gate profil dynamique *)
    WinchBrakeOpenDelayEffectiveS : REAL;             (* . [LOC] Delai ouverture applique apres gate profil dynamique *)
    WinchBrakeCloseDelayEffectiveS : REAL;            (* . [LOC] Delai fermeture applique apres gate profil dynamique *)
END_VAR

// === IMPLEMENTATION ===

{region "§1 Repli image reelle banc desactive"}
IF NOT Enable THEN
    // 🔌 Banc désactivé : repli sur l'image réelle, aucune simulation en cours
    KoboldMeasureEnablePrevious := FALSE;
    KoboldAutoEpisodeActive := FALSE;
    instKoboldPowerUpTimer(IN := FALSE);
    Ready       := FALSE;
    Busy        := FALSE;
    Done        := FALSE;
    Winch       := HwReal.Winch;
    Translation := HwReal.Translation;
    Operator    := HwReal.Operator;
    Machine     := HwReal.Machine;
    instSimJoystick(Enable := FALSE);
    RETURN;
END_IF;

// ▶️ Banc actif : le cycle de simulation démarre pour ce scan.
// 🔒 Le comptage brut M1/M2 (`_SimEncoderRawPosM1`/`M2`, GVL_PERSISTENT) n'est JAMAIS réécrit ici :
//    `FB_Sim_Encoder` en reste le producteur unique (accumulation signée / preset). L'origine de banc
//    plausible vient de l'initialisation DÉCLARÉE `GVL_PERSISTENT` (1 000 000 pts), pas d'une
//    réinjection conditionnelle : un 0 lu ici n'est PAS une mémoire vierge, c'est un point de passage
//    légitime du compteur SIGNÉ. Le banc ne réécrit donc aucune mémoire codeur, pas même pour
//    « initialiser » une valeur lue à 0 — une telle réinjection (1 100 000 pts = 268,55 m de position
//    publiée en un seul scan, sans mouvement ni défaut et référence de homing conservée)
//    transformerait un zéro réel en téléportation de position.
Ready := TRUE;
Busy  := TRUE;
Done  := FALSE;

{endregion}

{region "§2 Simulation treuils M1/M2"}
// ── 1. MODÈLE TREUILS (M1 + M2) ─────────────────────────────────────────────
// Presets codeurs : déclenchés si PresetTriggerCmd = 2
M1_PresetCmd := (M1_PresetTriggerCmd = 2);
M2_PresetCmd := (M2_PresetTriggerCmd = 2);
WinchSpeedReportTauEffectiveS := SEL(SimWinchDynamicsActive, 0.0, SimWinchSpeedReportTauS);
WinchBrakeOpenDelayEffectiveS := SEL(SimWinchDynamicsActive, 0.0, SimWinchBrakeOpenDelayS);
WinchBrakeCloseDelayEffectiveS := SEL(SimWinchDynamicsActive, 0.0, SimWinchBrakeCloseDelayS);

// Conversions d'injection d'écart synchro (0.5m -> points codeur avec 8192 pts/tour, 2m/tour)
// 1m = 4096 points codeur.
M1_OffsetPts := REAL_TO_DINT(SimSyncDeviationOffset_M * 4096.0);
M2_OffsetPts := REAL_TO_DINT(SimSyncDeviationOffset_M * 4096.0);

// Une plongée auto fige ses réglages avant l'arrêt : modifier l'IHM pendant AX5..AX8
// ne crée ni faux front fond ni changement de roulis en cours de mouvement.
IF KoboldMeasureEnable AND NOT KoboldMeasureEnablePrevious THEN
    KoboldAutoEpisodeActive := SimKoboldAutoModeActive;
    KoboldAutoDepthEpisode_M := SimKoboldAutoDepth_M;
    KoboldPowerUpEpisodeTime := SimKoboldPowerUpTime;
END_IF;
KoboldMeasureEnablePrevious := KoboldMeasureEnable;

// Instance modèle codeur M1
instSimEncoderM1(
    Enable              := TRUE,
    RelayFwd            := M1_RelayFwd,
    RelayRev            := M1_RelayRev,
    StepNumber          := M1_StepNumber,
    PresetCmd           := M1_PresetCmd,
    PresetValue         := M1_PresetValueOut,
    SpeedScaleFactor    := SimEncoderSpeedFactor,
    CoastDistanceM      := 0.0,
    SpeedReportTauS     := WinchSpeedReportTauEffectiveS,
    TestOffsetCmd       := SimSyncDeviationInjectM1,
    TestOffsetPts       := M1_OffsetPts,
    MechanicStopEngaged := FALSE,
    RawPos              := RawPosM1
);

// T317 exploratoire -- electrique+charge+couplage M1/M2, diagnostic seul (Winch.* metier deja
// consomme via M2_TensionedCable_DI ci-dessous). Couplage/charge cables sur stimuli de banc en
// attente des signaux reels amont (CoupledBoth, benne au sol) -- cf. registre PLAN_T317.
instWinchElectricalM1(
    Enable                := Enable AND SimWinchElectricalDiagnosticsActive,
    StepCmd               := MAX(1, M1_StepNumber),
    DirectionCmd          := SEL(M1_RelayRev, 1, -1),
    NetworkVoltageAct_V   := 400.0,
    LoadFrac_Ratio         := SEL(SimBucketJamActive, SimWinchLoadFrac_Ratio, CST_SimBucketJamLoadFrac_Ratio),
    IsBucketGrounded      := KoboldBottomTouchPrev_DI,
    IsCoupledToPeer        := SimWinchCoupledActive,
    PeerTorque_Nm          := PeerTorqueM2Prev_Nm,
    PeerSpeed_Rpm          := PeerSpeedM2Prev_Rpm
);
IF SimWinchElectricalDiagnosticsActive THEN
    MotorTorqueM1_Nm := instWinchElectricalM1.MotorTorque_Nm;
    MotorIsStalledM1 := instWinchElectricalM1.IsStalled;
    PeerTorqueM1Prev_Nm := instWinchElectricalM1.MotorTorque_Nm;
    PeerSpeedM1Prev_Rpm := instWinchElectricalM1.SpeedAct_Rpm;
ELSE
    MotorTorqueM1_Nm := 0.0;
    MotorIsStalledM1 := FALSE;
    PeerTorqueM1Prev_Nm := 0.0;
    PeerSpeedM1Prev_Rpm := 0.0;
END_IF;

instWinchElectricalM2(
    Enable                := Enable AND SimWinchElectricalDiagnosticsActive,
    StepCmd               := MAX(1, M2_StepNumber),
    DirectionCmd          := SEL(M2_RelayRev, 1, -1),
    NetworkVoltageAct_V   := 400.0,
    LoadFrac_Ratio         := SEL(SimBucketJamActive, SimWinchLoadFrac_Ratio, CST_SimBucketJamLoadFrac_Ratio),
    IsBucketGrounded      := KoboldBottomTouchPrev_DI,
    IsCoupledToPeer        := SimWinchCoupledActive,
    PeerTorque_Nm          := PeerTorqueM1Prev_Nm,
    PeerSpeed_Rpm          := PeerSpeedM1Prev_Rpm
);
IF SimWinchElectricalDiagnosticsActive THEN
    MotorTorqueM2_Nm := instWinchElectricalM2.MotorTorque_Nm;
    MotorIsStalledM2 := instWinchElectricalM2.IsStalled;
    PeerTorqueM2Prev_Nm := instWinchElectricalM2.MotorTorque_Nm;
    PeerSpeedM2Prev_Rpm := instWinchElectricalM2.SpeedAct_Rpm;
ELSE
    MotorTorqueM2_Nm := 0.0;
    MotorIsStalledM2 := FALSE;
    PeerTorqueM2Prev_Nm := 0.0;
    PeerSpeedM2Prev_Rpm := 0.0;
END_IF;

// Détection coupure relais M2 pour renouveler la dispersion pseudo-aléatoire (±0.1m)
IF (M2_RelayFwdPrev AND NOT M2_RelayFwd) OR (M2_RelayRevPrev AND NOT M2_RelayRev) THEN
    // Générateur LCG 32-bit standard : X_{n+1} = (1103515245 * X_n + 12345) MOD 2^31
    RandomSeed := (RandomSeed * 1103515245 + 12345) AND 16#7FFFFFFF;
    M2_EffectiveCoastM := (UDINT_TO_REAL(RandomSeed MOD 2000) / 10000.0) - 0.10;
END_IF;
M2_RelayFwdPrev := M2_RelayFwd;
M2_RelayRevPrev := M2_RelayRev;

// Manœuvre benne seule : M2 tourne, M1 est au repos (ouverture ou fermeture benne pure)
M2BucketOnlyActive := (M2_RelayFwd XOR M2_RelayRev) AND NOT M1_RelayFwd AND NOT M1_RelayRev;

// Descente conjointe physique (les deux treuils déroulent simultanément sous charge)
// Purement mécanique et basé sur les relais : AUCUNE dépendance à un mode ou au PRG_03.
M2CoupledDescentActive := SimM2CoupledDescentModelActive
                          AND M1_RelayRev AND M2_RelayRev
                          AND NOT M1_RelayFwd AND NOT M2_RelayFwd;

// Vitesses de palier nominales
SpeedM1_Mps := 0.2 + (INT_TO_REAL(MAX(M1_StepNumber, 1)) - 1.0) * 0.2;
SpeedM2_Mps := 0.2 + (INT_TO_REAL(MAX(M2_StepNumber, 1)) - 1.0) * 0.2;

// Facteur vitesse M2 :
// 1) En manœuvre benne seule : accélération via SimBucketSpeedFactor
// 2) En descente couplée benne ouverte : bridage de la vitesse de M2 à celle de M1 (zéro dérive -11m/-13m)
// 3) Nominal : SimEncoderSpeedFactor
M2EffectiveSpeedScaleFactor := SimEncoderSpeedFactor;
IF M2BucketOnlyActive THEN
    M2EffectiveSpeedScaleFactor := SimEncoderSpeedFactor * MAX(0.1, SimBucketSpeedFactor);
ELSIF M2CoupledDescentActive THEN
    // 🪝 Descente conjointe physique (M1 entraîné par la charge de benne, M2 freiné par réducteurs) :
    // M2 a un retard naturel proportionnel de 3% mesuré sur trace réelle (trace 36 : ~0.60 m à 20 m, ~1.5 m à 50 m).
    // Cela fait monter l\'écart (M2 - M1) progressivement et fidèlement avec la profondeur, quel que soit le mode (MANU/AUTO).
    IF SpeedM2_Mps > 0.01 THEN
        M2EffectiveSpeedScaleFactor := SimEncoderSpeedFactor * (SpeedM1_Mps / SpeedM2_Mps) * 0.97;
    ELSE
        M2EffectiveSpeedScaleFactor := SimEncoderSpeedFactor * MAX(0.0, SimM2CoupledDescentFactor);
    END_IF;
END_IF;

// P02 consomme la mesure publiée au scan précédent. Reconstituer le déplacement
// de ce scan évite un trou d'un cycle lors du seuil d'arrêt de FB_Bucket.
M2ExpectedStepDistance_M := (1.0 + (INT_TO_REAL(MAX(M2_StepNumber, 1)) - 1.0) * 0.25)
                            * MAX(0.0, M2EffectiveSpeedScaleFactor)
                            * CST_SimBenchCycleTimeS;
M2OpenStopThreshold_M := BucketOffsetOpen_M + MAX(0.0, BucketOpenAnticipation_M)
                         + M2ExpectedStepDistance_M;

// Armer le roulis long uniquement à l'approche du seuil d'ouverture AX15B.
// Un jog manuel, un homing ou un arrêt ailleurs garde le roulis historique.
IF NOT M2_RelayRev OR M2_RelayFwd THEN
    M2AutoOpenCoastArmed := FALSE;
ELSIF SimWinchCouplingModelActive AND BucketAx15bOpenActive
      AND NOT M1_RelayFwd AND NOT M1_RelayRev
      AND (M2_CablePos_M - M1_CablePos_M)
          <= M2OpenStopThreshold_M THEN
    M2AutoOpenCoastArmed := TRUE;
END_IF;

// À l'arrêt anticipé automatique, le roulis couvre seulement l'écart restant
// jusqu'à la butée ouverte : il ne sur-ouvre pas et ne modifie pas le jog manuel.
M2EffectiveCoastDistance_M := M2_EffectiveCoastM;
IF M2AutoOpenCoastArmed THEN
    M2OpenDistanceRemaining_M := MAX(0.0, M2_CablePos_M - M1_CablePos_M
                                          - BucketOffsetOpen_M - M2ExpectedStepDistance_M);
    M2EffectiveCoastDistance_M := MIN(MAX(0.0, BucketOpenAnticipation_M),
                                      M2OpenDistanceRemaining_M);
END_IF;

// Butée mécanique benne (T421) : bloque le mouvement de manœuvre benne à la butée.
// N'arrête M2 que s'il est commandé SEUL vers la butée (ouverture sous BucketOffsetOpen_M
// ou fermeture au-dessus de BucketOffsetCloseM).
M2_MechanicStopEngaged := SimWinchCouplingModelActive
                          AND WinchesHomed
                          AND (((M2_CablePos_M - M1_CablePos_M) <= (BucketOffsetOpen_M - 0.40) AND M2_RelayRev AND NOT M1_RelayRev)
                               OR ((M2_CablePos_M - M1_CablePos_M) >= BucketOffsetCloseM AND M2_RelayFwd AND NOT M1_RelayFwd));

// Instance modèle codeur M2 (dynamique T421 continue, CoastDistanceM=0)
instSimEncoderM2(
    Enable              := TRUE,
    RelayFwd            := M2_RelayFwd,
    RelayRev            := M2_RelayRev,
    StepNumber          := M2_StepNumber,
    PresetCmd           := M2_PresetCmd,
    PresetValue         := M2_PresetValueOut,
    SpeedScaleFactor    := M2EffectiveSpeedScaleFactor,
    CoastDistanceM      := 0.0,
    SpeedReportTauS     := WinchSpeedReportTauEffectiveS,
    TestOffsetCmd       := SimSyncDeviationInjectM2,
    TestOffsetPts       := M2_OffsetPts,
    MechanicStopEngaged := M2_MechanicStopEngaged,
    RawPos              := RawPosM2
);

// L'épisode Kobold ne produit que la DI. Le cycle commande l'arrêt ; les FB codeurs
// conservent leur roulis historique après la retombée des relais.
IF NOT KoboldMeasureEnable AND NOT M1_RelayRev AND NOT M2_RelayRev
   AND NOT M1_RelayFwd AND NOT M2_RelayFwd THEN
    KoboldAutoEpisodeActive := FALSE;
END_IF;

// Recopie structures Winch simulées :
// 🛑 POLARITÉ DE FREIN SIMULÉ : 1 = contacteur commandé = frein OUVERT.
// Câblage réel : DI = 1 ⟺ frein OUVERT. Le modèle produit donc M1_BrakeIsOpen_DI := M1_BrakeCmd !
// Delai electrique/meca opt-in : SimWinchBrakeOpenDelayS/CloseDelayS=0.0 -> bascule le
// meme scan (comportement historique inchange, TC-P13-012). >0 -> retour retarde, sans jamais
// inverser la polarite (M1_BrakeIsOpenState suit toujours M1_BrakeCmd, juste avec latence).
IF M1_BrakeCmd THEN
    IF NOT M1_BrakeIsOpenState THEN
        M1_BrakeOpenTimerS := M1_BrakeOpenTimerS + CST_SimBenchCycleTimeS;
        IF M1_BrakeOpenTimerS >= MAX(0.0, WinchBrakeOpenDelayEffectiveS) THEN
            M1_BrakeIsOpenState := TRUE;
            M1_BrakeOpenTimerS := 0.0;
        END_IF;
    END_IF;
    M1_BrakeCloseTimerS := 0.0;
ELSE
    IF M1_BrakeIsOpenState THEN
        M1_BrakeCloseTimerS := M1_BrakeCloseTimerS + CST_SimBenchCycleTimeS;
        IF M1_BrakeCloseTimerS >= MAX(0.0, WinchBrakeCloseDelayEffectiveS) THEN
            M1_BrakeIsOpenState := FALSE;
            M1_BrakeCloseTimerS := 0.0;
        END_IF;
    END_IF;
    M1_BrakeOpenTimerS := 0.0;
END_IF;
Winch.M1_BrakeIsOpen_DI        := M1_BrakeIsOpenState;
// Retour UNIQUE « tous contacteurs retombés » = sens ET vitesse.
// Omettre les paliers ferait croire à l'arrêt pendant les transitoires → Méca A armée à tort.
Winch.M1_ContactorsReleased_DI := NOT (M1_RelayFwd OR M1_RelayRev
                                    OR M1_SpeedContactor_1 OR M1_SpeedContactor_2
                                    OR M1_SpeedContactor_3 OR M1_SpeedContactor_4);
Winch.M1_ThermalOk_DI          := TRUE; // Sauf panne simulée

IF M2_BrakeCmd THEN
    IF NOT M2_BrakeIsOpenState THEN
        M2_BrakeOpenTimerS := M2_BrakeOpenTimerS + CST_SimBenchCycleTimeS;
        IF M2_BrakeOpenTimerS >= MAX(0.0, WinchBrakeOpenDelayEffectiveS) THEN
            M2_BrakeIsOpenState := TRUE;
            M2_BrakeOpenTimerS := 0.0;
        END_IF;
    END_IF;
    M2_BrakeCloseTimerS := 0.0;
ELSE
    IF M2_BrakeIsOpenState THEN
        M2_BrakeCloseTimerS := M2_BrakeCloseTimerS + CST_SimBenchCycleTimeS;
        IF M2_BrakeCloseTimerS >= MAX(0.0, WinchBrakeCloseDelayEffectiveS) THEN
            M2_BrakeIsOpenState := FALSE;
            M2_BrakeCloseTimerS := 0.0;
        END_IF;
    END_IF;
    M2_BrakeOpenTimerS := 0.0;
END_IF;
Winch.M2_BrakeIsOpen_DI        := M2_BrakeIsOpenState;
Winch.M2_ContactorsReleased_DI := NOT (M2_RelayFwd OR M2_RelayRev
                                    OR M2_SpeedContactor_1 OR M2_SpeedContactor_2
                                    OR M2_SpeedContactor_3 OR M2_SpeedContactor_4);
Winch.M2_ThermalOk_DI          := TRUE;

// Cohérent avec M2_TensionedCable_DI (sain par défaut) : capteur TOP libre en simu,
// sauf stimulus manuel SimTopPositionActive (injection de fait capteur au banc).
Winch.M1M2_TopPositionFree_DI  := NOT SimTopPositionActive;
// Le Kobold ne deduit pas l'etat cable : seul le stimulus safety explicite injecte une panne.
Winch.M2_TensionedCable_DI     := NOT SimM2TensionedCableFaultInject;

Winch.COD1_PosValue            := instSimEncoderM1.RawPosOut;
Winch.COD1_SpdValue            := instSimEncoderM1.RawSpdOut;
Winch.COD1_Alarms              := 0;
Winch.COD1_Warnings            := 0;
Winch.COD1_DeviceState         := DEVICE_STATE.RUNNING; // État device RUNNING (bus OK)

Winch.COD2_PosValue            := instSimEncoderM2.RawPosOut;
Winch.COD2_SpdValue            := instSimEncoderM2.RawSpdOut;
Winch.COD2_Alarms              := 0;
Winch.COD2_Warnings            := 0;
Winch.COD2_DeviceState         := DEVICE_STATE.RUNNING; // État device RUNNING

{region "§2bis Rattrapage mecanique M1/M2"}
// La benne relie mecaniquement les deux treuils. En MONTEE couplee et sans blocage, le jeu relatif
// est repris : Delta = PosM2 - PosM1 rejoint la BUTEE mecanique benne FERMEE (OffsetCloseM).
// Sans ce rattrapage, un ecart residuel (trou metier de fermeture : coupure d'anticipation a 13,8 m
// alors que l'etat ferme exige 14,0 m) laisse la benne "non fermee" et plafonne la montee au palier 1.
// 🔒 Le modele n'ecrit QUE l'image publiee (Winch.COD2_PosValue) -- JAMAIS RawPosM2, memoire
//    persistante du codeur dont FB_Sim_Encoder reste l'unique producteur.
// 🔒 MONTEE UNIQUEMENT : la descente couplee reste au modele existant SimM2CoupledDescentModelActive
//    (exclusion mutuelle : les deux modeles ne s'appliquent jamais ensemble).
// 🔒 Cible = BUTEE MECANIQUE benne fermee (BucketOffsetCloseM) : seule valeur qui fasse converger
//    l'ouverture benne vers 0 % ; une cible intermediaire laisse un ecart plancher jamais
//    corrigible. Le sens unique (correction seulement si Delta < cible) et le bornage de pente
//    (LIMIT + MIN(cible - Delta)) interdisent tout depassement de butee.
WinchCouplingBothSameDir := (M1_RelayFwd AND M2_RelayFwd) OR (M1_RelayRev AND M2_RelayRev);
WinchCouplingGate := SimWinchCouplingModelActive
                     AND WinchCouplingBothSameDir
                     AND M1_RelayFwd AND NOT M1_RelayRev        // montee uniquement
                     AND M1_BrakeIsOpenState AND M2_BrakeIsOpenState
                     AND Winch.M2_TensionedCable_DI            // cable tendu : sinon aucun effort transmis
                     AND NOT KoboldBottomTouchPrev_DI          // benne au fond : aucun mouvement reel
                     AND NOT (M1_PresetCmd OR M2_PresetCmd)    // jamais pendant un preset/homing
                     AND NOT SimBucketJamActive;               // mâchoires bloquees : aucun rattrapage
WinchCouplingActive := WinchCouplingGate;
WinchCouplingCorrectionPts := 0;
IF WinchCouplingGate THEN
    WinchCouplingDelta_M := M2_CablePos_M - M1_CablePos_M;
    // Cible = butee mecanique benne FERMEE (ecart relatif 0 %). Le sens unique et le bornage
    // de pente garantissent qu'aucune correction ne depasse cette butee.
    WinchCouplingTarget_M := BucketOffsetCloseM;
    IF WinchCouplingDelta_M < WinchCouplingTarget_M THEN
        WinchCouplingCorrection_M := (WinchCouplingTarget_M - WinchCouplingDelta_M)
                                     * CST_SimBenchCycleTimeS
                                     / (CST_SimWinchCouplingTauS + CST_SimBenchCycleTimeS);
        // Sens unique + bornage (§6) : jamais de saut, jamais au-dela de la cible
        WinchCouplingCorrection_M := LIMIT(0.0, WinchCouplingCorrection_M,
                                           MIN(CST_SimWinchCouplingStepMax_M,
                                               WinchCouplingTarget_M - WinchCouplingDelta_M));
        WinchCouplingCorrectionDInt := REAL_TO_DINT(WinchCouplingCorrection_M
                                                    * CST_SimWinchCouplingPtsPerM);
        IF WinchCouplingCorrectionDInt > 0 THEN
            WinchCouplingAccumPts := WinchCouplingAccumPts + WinchCouplingCorrectionDInt;
            WinchCouplingCorrectionPts := WinchCouplingCorrectionDInt;
        END_IF;
    END_IF;
ELSIF M2_RelayRev AND NOT M2_RelayFwd THEN
    // Ouverture commandee : la reprise de jeu est relachee (le cable de fermeture devide),
    // sinon l'image M2 masquerait l'ouverture reelle.
    WinchCouplingCorrectionDInt := REAL_TO_DINT(CST_SimWinchCouplingStepMax_M
                                                * CST_SimWinchCouplingPtsPerM);
    WinchCouplingAccumPts := MAX(0, WinchCouplingAccumPts - WinchCouplingCorrectionDInt);
END_IF;
// Un preset/homing rend la reference absolue : l'offset de reprise de jeu n'a plus de sens.
IF M1_PresetCmd OR M2_PresetCmd THEN
    WinchCouplingAccumPts := 0;
END_IF;
// Report sur l'IMAGE uniquement (le raw persistant n'est jamais touche), et seulement quand le
// modele est actif : en mode desactive, l'image reste strictement celle du codeur.
IF SimWinchCouplingModelActive AND (WinchCouplingAccumPts > 0) THEN
    Winch.COD2_PosValue := Winch.COD2_PosValue + DINT_TO_UDINT(WinchCouplingAccumPts);
END_IF;
{endregion}

{endregion}

{region "§3 Simulation translation M3"}
// ── 2. MODÈLE TRANSLATION M3 (AC600) ─────────────────────────────────────────
M3_RelayFwd := M3_ReqTremie AND NOT M3_ReqMaintenance;
M3_RelayRev := M3_ReqMaintenance AND NOT M3_ReqTremie;

instSimTranslation(
    Enable          := TRUE,
    ReqTremie       := M3_RelayFwd,
    ReqMaintenance  := M3_RelayRev,
    SpeedTgt_Pct    := M3_SpeedCmd_Pct,
    PosTremie_M        := M3_PosTremie_M,
    PosPV_M            := M3_PosPV_M,
    PosP2_M            := M3_PosP2_M,
    PosP1_M            := M3_PosP1_M,
    PosMaintenance_M   := M3_PosMaintenance_M,
    GainMetersPerHzSec := M3_OdometryGain,
    EndStopMargin_M    := SimM3EndStopMargin_M,
    MaxFreq_Hz      := CST_M3MaxFreq_Hz,
    SpeedFactor     := SimM3SpeedFactor,
    BrakeReleaseCmd := M3_BrakeCmd,
    SensorIntermittenceActive := SimM3SensorIntermittenceActive,
    SensorStabilizationS := SimM3SensorStabilizationS,
    SensorElectricalDelayS := SimM3SensorElectricalDelayS,
    SensorIntermittencePeriodS := SimM3SensorIntermittencePeriodS,
    SensorHysteresis_M := SimM3SensorHysteresis_M,
    SensorLoadAngleTriggerRad := SimM3SensorLoadAngleTriggerRad,
    SensorScenarioSeed := SimM3SensorScenarioSeed,
    SensorBlipTransitions := SimM3SensorBlipTransitions,
    SensorBlipDurationS := SimM3SensorBlipDurationS,
    BrakeFaultCloseWhileRunning := SimM3BrakeFaultCloseWhileRunning,
    BrakeFaultCloseDelay_S := SimM3BrakeFaultCloseDelayS,
    EndStopRecoilMax_M := SimM3EndStopRecoilMax_M,
    LoadReactionGain_Mps2 := SimM3LoadReactionGain_Mps2,
    BrakePhysicalActive := SimM3BrakePhysicalActive,
    BrakeDecel_Mps2 := SimM3BrakeDecel_Mps2,
    CartFreeActive := SimM3CartFreeActive,
    LoadMassRatio := SimM3LoadMassRatio,
    RollingFriction_Mps2 := SimM3RollingFriction_Mps2,
    Slope_Mps2 := SimM3Slope_Mps2,
    SensorCamDropoutActive := SimM3SensorCamDropoutActive,
    SensorCamDropoutStart_M := SimM3SensorCamDropoutStart_M,
    SensorCamDropoutWidth_M := SimM3SensorCamDropoutWidth_M
);
M3BrakeFaultCloseActive := instSimTranslation.BrakeFaultCloseActive;
M3SensorBlipActive := instSimTranslation.SensorBlipActive;
M3ObsPositionTrue_M := instSimTranslation.PositionTrue_M;
M3ObsPositionError_M := instSimTranslation.PositionTrue_M - M3_EstimatedPos_M;
M3ObsOvershootLast_M := instSimTranslation.ObsOvershootLast_M;
M3ObsOvershootSensorId := instSimTranslation.ObsOvershootSensorId;
M3ObsEndStopHitCount := instSimTranslation.ObsEndStopHitCount;
M3ObsEndStopImpactSpeed_Mps := instSimTranslation.ObsEndStopImpactSpeed_Mps;
M3ObsBrakeClosedMovingCount := instSimTranslation.ObsBrakeClosedMovingCount;
M3ObsCartFree := instSimTranslation.ObsCartFree;
M3ObsFreeRollLast_M := instSimTranslation.ObsFreeRollLast_M;

// Remplissage capteurs de position M3 : l'override manuel conserve exactement le
// même ordre que FB_Translation_PositionDecoder (bit4=Trémie ... bit0=Maintenance).
IF SimM3SensorsWordOverrideActive THEN
    Translation.M3_PosTremie_DI      := SimM3SensorsWord.4;
    Translation.M3_PosPV_DI          := SimM3SensorsWord.3;
    Translation.M3_PosPVP2_DI        := SimM3SensorsWord.2;
    Translation.M3_PosP1_DI          := SimM3SensorsWord.1;
    Translation.M3_PosMaintenance_DI := SimM3SensorsWord.0;
ELSE
    Translation.M3_PosTremie_DI      := instSimTranslation.PosTremie;
    Translation.M3_PosPV_DI          := instSimTranslation.PosPV;
    Translation.M3_PosPVP2_DI        := instSimTranslation.PosP2;
    Translation.M3_PosP1_DI          := instSimTranslation.PosP1;
    Translation.M3_PosMaintenance_DI := instSimTranslation.PosMaintenance;
END_IF;

// Retour auxiliaire du frein, distinct de la commande electrique.
Translation.M3_BrakeIsOpen_DI    := instSimTranslation.BrakeContactOpen;

// Thermique moteur/variateur AC600 — pas de panne simulée, toujours OK (comme Winch.M1/M2_ThermalOk_DI)
Translation.M3_ThermalOK_DI      := TRUE;

// Simulation StatusWord AC600 : Bit 0 (Power Ready) = 1, Bit 7 (Comm Ready) = 1 -> 16#0087 en mouvement
// Bit0 retombe à l'arrêt, cohérent avec un variateur qui confirme l'arrêt sans rester "actif" —
// FB_Safety_Translation lit ce bit comme indicateur "mouvement non commandé" (Méca B, TonMecaB 3s) :
// un Bit0 forcé à 1 en continu à l'arrêt déclencherait un PowerCutOff simulé permanent après 3s.
// DrivePowerReady (diagnostic IHM seul, non consommé par un interlock) est le seul autre lecteur,
// aucune régression de mouvement possible.
IF instSimTranslation.ActualFrequency_Hz > 0.5 THEN
    M3_StatusWordSim := 16#0087; // + Operating/Running
ELSE
    M3_StatusWordSim := 16#0080; // Comm Ready seul -- Bit0 retombé, arrêt confirmé
END_IF;
M3_ActualFreqHz := REAL_TO_UINT(LIMIT(0.0, instSimTranslation.ActualFrequency_Hz, CST_M3MaxFreq_Hz) * 100.0);

Translation.M3_StatusWord        := M3_StatusWordSim;
Translation.M3_ActualFrequencyHz := M3_ActualFreqHz;
Translation.AC600_DeviceState    := DEVICE_STATE.RUNNING; // État device RUNNING

{endregion}

{region "§4 Simulation operateur joystick"}
// ── 3. MODÈLE OPÉRATEUR / JOYSTICK ───────────────────────────────────────────
IF NOT OperatorSourceActive THEN
    // Le geste ne continue pas en arriere-plan lorsque le domaine est reel.
    instSimJoystick(Enable := FALSE);
    Operator := HwReal.Operator;
ELSE
    SimJoystickManualNeutral := (SimJoystickRawX = 5000) AND (SimJoystickRawY = 5000);
    SimJoystickGesturePermit := SimJoystickManualNeutral AND NOT SimJoystickRawButton;
    instSimJoystick(
        Enable              := TRUE,
        GesturePermit       := SimJoystickGesturePermit,
        NeutralRaw          := 5000,
        MaxRaw              := 10000,
        BtnLeft_Rev_TREMIE  := SimJoystickLeft_Rev_TREMIE_Active,
        BtnRight_Fwd_MAINT  := SimJoystickRight_Fwd_MAINT_Active,
        BtnFwd_Up_Close     := SimJoystickFwd_Up_Close_Active,
        BtnRev_Down_Open    := SimJoystickRev_Down_Open_Active,
        OvershootActive     := SimJoystickOvershoot_Active,
        BagotementActive    := SimJoystickBagotement_Active,
        CycleTimeS          := 0.010
    );

    // Une seule source possede les trois signaux : aucun melange bouton/axes.
    // La propriete automatique persiste au retour et si un stimulus manuel est en conflit.
    IF instSimJoystick.ModelActive THEN
        Operator.JoyXRaw_ANA1 := instSimJoystick.RawX;
        Operator.JoyYRaw_ANA2 := instSimJoystick.RawY;
        Operator.JoyBtnRaw := instSimJoystick.RawButton;
    ELSE
        // Modèle au repos → stimulus analogique avancé (mode « sans bouton »).
        Operator.JoyXRaw_ANA1 := SimJoystickRawX;
        Operator.JoyYRaw_ANA2 := SimJoystickRawY;
        Operator.JoyBtnRaw := SimJoystickRawButton;
    END_IF;

    Operator.CanBusState      := 2; // CANbusState 2 = ACTIVE
    Operator.JOY1_DeviceState := DEVICE_STATE.RUNNING; // État device RUNNING
END_IF;

{endregion}

{region "§5 Simulation securite et image machine"}
// ── 4. MODÈLE SÉCURITÉ & COMMUNS MACHINE ─────────────────────────────────────
instSimSafety(
    Enable            := TRUE,
    SimChainOkBit     := SimChainOkBit,
    SimPhaseRotationOkBit := SimPhaseRotationOkBit,
    PowerCutOff_A     := PowerKeepAlive_A,
    PowerCutOff_B     := PowerKeepAlive_B,
    PowerCutOffRequest:= PowerCutOffRequest,
    EmergencyArming   := EmergencyArming_RQ,
    BtnEmergencyStop  := BtnEmergencyStop,
    TestCutActive     := TestCutActive
);

Machine.PowerContactorEngaged_DI   := instSimSafety.SimContactorOk;
Machine.EmergencyChainClosed_DI    := instSimSafety.SimChainOk;
Machine.PhaseRotationOk_DI          := instSimSafety.SimPhaseRotationOk;
Machine.M1_M2_M3_BrakeThermalOk_DI     := TRUE;
instKoboldPowerUpTimer(IN := KoboldAutoEpisodeActive AND KoboldMeasureEnable
                        AND (M1_CablePos_M > KoboldAutoDepthEpisode_M),
                        PT := KoboldPowerUpEpisodeTime);
IF KoboldAutoEpisodeActive THEN
    Machine.M1_M2_KoboldBottomTouch_DI := instKoboldPowerUpTimer.Q
                                           AND (M1_CablePos_M > KoboldAutoDepthEpisode_M);
ELSE
    Machine.M1_M2_KoboldBottomTouch_DI := SimKoboldContactValue;
END_IF;
// T317 : memorise pour le prochain scan -- reutilise le VRAI capteur fond (Kobold), pas un
// stimulus invente, cf. retour utilisateur 2026-09-18 (le capteur fond existe deja reel+sim).
KoboldBottomTouchPrev_DI := Machine.M1_M2_KoboldBottomTouch_DI;
Machine.HydraulicThermalOk_DI          := TRUE;
Machine.TremieFull_OR_GateRaised_DI    := FALSE; // Pas encore câblé, simulé inactif par défaut

// ✅ Cycle de simulation terminé : les 4 images sont publiées pour ce scan
Busy := FALSE;
Done := TRUE;

{endregion}

END_FUNCTION_BLOCK
